Staubli VAL3: default.dtx


